FUNCTION_BLOCK T_SafeDecouple_Tests EXTENDS TcUnit.FB_TestSuite
VAR
    // Test_InputsLoopedToOutputsOnlyWhenRunning
    group_1 : T_SafeGroup;
    fb_1 : T_SafeDecouple(group := group_1);
END_VAR

Test_InputsLoopedToOutputsOnlyWhenRunning();

METHOD PRIVATE Test_InputsLoopedToOutputsOnlyWhenRunning
TcUnit.TEST(__POUNAME());
// act
group_1(Run := TRUE);
fb_1(DecIn3 := TRUE);
// assert
AssertEquals_BOOL(Expected := TRUE, Actual := fb_1.DecOut3, Message := 'input looped to output');
group_1(Run := FALSE);
fb_1(DecIn3 := TRUE);
AssertEquals_BOOL(Expected := FALSE, Actual := fb_1.DecOut3, Message := 'output off while the group is stopped');
TEST_FINISHED_NAMED(__POUNAME());
END_METHOD

END_FUNCTION_BLOCK

(* stored: Version 1.1.0.1
   POU T_SafeDecouple_Tests: Id {53c8a3f7-118d-5f6f-8073-5da89a3cdba1}, SpecialFunc None
   Method Test_InputsLoopedToOutputsOnlyWhenRunning: Id {a98a7e9d-5d5b-57af-a460-345e5764e19b} *)
